//---------------------------------------------------------------------------------------------------------------
//
//  HAUD 2026.11.07
//
//  - TowerControl - fb_DisposableHeros
//
//    - this class is nothing more than the handshake sequence and a timer
//
//    - the station bitmask is written for each production cycle
//      - ticketing involves a DistributorByTicket and its companion ProcessByTicket
//      - this mock up takes care of both tickets.
//        - Why do you need to send 2 tickets?
//          - Distributor and Process instance do not know each other (and this is on purpose to keep things loose and avoid thight coupling by design)
//            --> sending tickets should be done from one place only, so a Distributor sending a ticket internally to its Process would break that rule.
//            --> The Ticket transports the information about where the movers were sent to
//              --> The Process now needs to be told which stations to activate, the rest is ruled by the bitmask from the ticket. 
//
//    - top level transport abstractions are handshaked here:
//    --------------------------------------------
//    - top level transport abstractions
//      - Instances contain the required transport logic
//      - Instances control their assigned ProcessCollector
//      - Instances are controlled in timer based application
//
//
//---------------------------------------------------------------------------------------------------------------
FUNCTION_BLOCK fb_DisposableHeros // Soldier boy, made of clay, now an empty shell
VAR_INPUT
  Start         : BOOL;           // Back to the front
  DwellTime     : TIME;           // Sounding of the clock that ticks
  StationMask   : T_PROCESS;      // molded day by day
END_VAR
VAR
  // process index
  _nProcess               : E_INSTANCE; // whoami
  _nProcessConnect        : e_instance; // to whom am I connected? this is an idea to manage the two tickets for Distributor and Process
  _nProcessConnectTarget  : e_instance; // what is the target of the process to whom I am connected

  _stInstanceCtrl         : REFERENCE TO ARRAY[1..MAX_PROCESS] OF ST_INSTANCE_CTRL;
  _stInstanceState        : REFERENCE TO ARRAY[1..MAX_PROCESS] OF ST_INSTANCE_STATE;

  _wActivateStation       : T_PROCESS;
  _stProcessData          : ST_PROCESS_DATA;

  _ItfTicketList          : I_Process_LinkedList;
  _WriteResult            : ST_PROCESS_LIST_RESULT;

  _nState                 : UINT;
  _tonProcess             : Tc2_Standard.TON;

  _nTicketCount           : UDINT;  // since this is a mock up, there is no-one to clean this up
  _nTicketCountLimit      : UDINT;  // if <> 0 --> limit is active

  _tdx                    : UINT;
END_VAR

//---------------------------------------------------------------------------------------------------------------
//---------------------------------------------------------------------------------------------------------------
// CHECK() ??
// !! this is mock up code, there is no check
//
//---------------------------------------------------------------------------------------------------------------
//---------------------------------------------------------------------------------------------------------------
IF NOT Start THEN _nState   := 0; END_IF
//---------------------------------------------------------------------------------------------------------------
CASE _nState OF
  0:
    IF Start
    THEN
      _nState               := 10;
    END_IF

  10:
    CASE _stInstanceState[_nProcess].ProcessState
    OF
      E_INSTANCE_STATE.DISABLED:
        _stInstanceCtrl[_nProcess].Cmd        := E_INSTANCE_CMD.ENABLE;
        IF (_nProcessConnect > e_instance.INSTANCE_NULL)
        THEN
          memset(ADR(_stProcessData), 0, SIZEOF(_stProcessData));
          _nState                             := 20;
          _wActivateStation                   := StationMask; // this one is important, must be double checked before sending
        END_IF

      E_INSTANCE_STATE.ENABLED:
        CASE _stInstanceState[_nProcess].ProcessProgress
        OF
          E_PROGRESS.PROGRESS_OCCUPIED:       // allow infeed movement
            _tonProcess(IN := FALSE, 
                        PT := DwellTime);

            _stInstanceCtrl[_nProcess].Cmd    := E_INSTANCE_CMD.PROCEED;
        END_CASE

      E_INSTANCE_STATE.WORKING:               // this is for the ProcessByTicket standstill handshake
        CASE _stInstanceState[_nProcess].ProcessProgress
        OF
          E_PROGRESS.PROGRESS_BUSY:           // now every mover has arrived.
            _tonProcess(IN := TRUE, 
                        PT := DwellTime);

            IF (_tonProcess.Q)
            THEN
              memset(ADR(_stProcessData), 0, SIZEOF(_stProcessData));
              _stInstanceCtrl[_nProcess].Cmd := E_INSTANCE_CMD.WORK;
            END_IF

          E_PROGRESS.PROGRESS_OCCUPIED:       // time is fleeting
            _stInstanceCtrl[_nProcess].Cmd  := E_INSTANCE_CMD.FINISH;
        END_CASE

      E_INSTANCE_STATE.FINISH:                // madness takes its toll
        CASE _stInstanceState[_nProcess].ProcessProgress
        OF
          E_PROGRESS.PROGRESS_DONE:
            _tonProcess(IN := FALSE, 
                        PT := DwellTime);

            _stInstanceCtrl[_nProcess].Cmd    := E_INSTANCE_CMD.DISABLE;

            IF (_nProcessConnect > e_instance.INSTANCE_NULL)
            THEN
              memset(ADR(_stProcessData), 0, SIZEOF(_stProcessData));
              _nState                         := 30;
              _wActivateStation               := StationMask; // this one is important, must be double checked before sending
            END_IF
        END_CASE
    END_CASE
END_CASE
CASE _nState OF
  20:
    _nState                                   :=  10;
    TruncMask();

  30:
    _nState                                   := 100;
    TruncMask();
END_CASE
CASE _nState OF

  100:
    //-----------------------------------------------------------------------------  
    // the tickets
    //-----------------------------------------------------------------------------
    // first send the ticket to the Distributor
    _WriteResult                          := _ItfTicketList.AddTailValue(_stProcessData);
    // second write the ticket for the Process
    _stProcessData.nProcessId             := _nProcessConnect;
    _stProcessData.nTargetId              := _nProcessConnectTarget;
    // third send the ticket to the Process
    _WriteResult                          := _ItfTicketList.AddTailValue(_stProcessData);
    //-----------------------------------------------------------------------------
    _nTicketCount                         := _nTicketCount + 1;;
    //-----------------------------------------------------------------------------
    _nState                               := 1000;
END_CASE
CASE _nState OF

  1000:
    IF NOT (_nTicketCountLimit > 0)
    THEN
      _nState                             := 0;
    ELSE
      IF (_nTicketCount < _nTicketCountLimit)
      THEN
        _nState                           := 0;
      END_IF
    END_IF
END_CASE

METHOD PUBLIC BitGet : BOOL
VAR_INPUT
  inVal   : T_PROCESS;
  bitNo   : DINT;
END_VAR
VAR
  wConst : T_PROCESS := 1;
END_VAR
IF ( inVal AND SHL( wConst,TO_SINT(bitNo) MOD TO_INT(SIZEOF(T_PROCESS)*8) ) ) > 0
THEN
  BitGet := TRUE;
ELSE
  BitGet := FALSE;
END_IF
END_METHOD

METHOD PUBLIC BitSet : T_PROCESS
VAR_INPUT
  inVal   : T_PROCESS;
  bitNo   : DINT;
END_VAR
VAR
  wConst  : T_PROCESS := 1;
END_VAR
BitSet := inVal OR SHL( wConst,TO_SINT(bitNo) MOD TO_INT(SIZEOF(T_PROCESS)*8) );
END_METHOD

PROPERTY InstanceCtrl : REFERENCE TO ARRAY[1..MAX_PROCESS] OF ST_INSTANCE_CTRL
SET
_stInstanceCtrl ref= InstanceCtrl;
END_SET
END_PROPERTY

PROPERTY InstanceState : REFERENCE TO ARRAY[1..MAX_PROCESS] OF ST_INSTANCE_STATE
SET
_stInstanceState ref= InstanceState;
END_SET
END_PROPERTY

PROPERTY ProcessId : E_INSTANCE
GET
ProcessId := _nProcess;
END_GET
SET
_nProcess := ProcessId;
END_SET
END_PROPERTY

PROPERTY ProcessId_Connect : E_INSTANCE
GET
ProcessId_Connect := _nProcessConnect;
END_GET
SET
_nProcessConnect := ProcessId_Connect;
END_SET
END_PROPERTY

PROPERTY ProcessId_ConnectTarget : E_INSTANCE
GET
ProcessId_ConnectTarget := _nProcessConnectTarget;
END_GET
SET
_nProcessConnectTarget := ProcessId_ConnectTarget;
END_SET
END_PROPERTY

PROPERTY TicketLinkedList : I_Process_LinkedList
SET
_ItfTicketList := TicketLinkedList;
END_SET
END_PROPERTY

METHOD TruncMask : BOOL
VAR_INPUT
END_VAR
// transfer station mask only in the range possible to handle in connected process (StationCount)
_stProcessData.nProcessId                 := _nProcess;
_stProcessData.nTargetId                  := _nProcessConnect;

FOR _tdx := 1 TO _stInstanceState[_nProcessConnect].StationCount
DO
  IF (BitGet(_wActivateStation, _tdx-1))
  THEN
    _stProcessData.wTarget                := BitSet(_stProcessData.wTarget, _tdx-1);
  END_IF      
END_FOR

TruncMask := TRUE;
END_METHOD

END_FUNCTION_BLOCK

(* stored: Version 1.1.0.1
   POU fb_DisposableHeros: Id {57ff81e0-db35-4988-adb1-755f5d46de47}, SpecialFunc None
   Method BitGet: Id {57c98de9-b3fd-4f7e-920b-502f6210a0a0}
   Method BitSet: Id {075d513b-2170-4aca-a2e9-2a16152dac6f}
   Property InstanceCtrl: Id {3363ce1e-638f-4a56-a7d9-502d7b3ac384}
   Set Set: Id {f01b16e3-e7c7-4d66-96b7-a5ce7482bb16}
   Property InstanceState: Id {4aad0611-ac13-4ac9-9913-e5032aa8988a}
   Set Set: Id {d6f80117-bb3a-400d-a886-057ce4f9cae4}
   Property ProcessId: Id {b0d1a924-6241-4335-be39-966d3f9b0719}
   Get Get: Id {4b563e78-35ca-46fa-a429-91bad99e170e}
   Set Set: Id {566aa5ef-d2c9-4a5c-8d5d-3fca3942f3dd}
   Property ProcessId_Connect: Id {abcc06e1-efe7-4aa9-9516-be1588519f38}
   Get Get: Id {b63ddabd-1e94-4d54-b9cd-0e5cfc49b660}
   Set Set: Id {97104ab0-4bc8-47e4-aa6e-413c64ff8466}
   Property ProcessId_ConnectTarget: Id {da385cf2-47a3-4307-bcdb-9af574222ed1}
   Get Get: Id {e9f241da-b82b-4801-b1f0-50eb7bef7352}
   Set Set: Id {95ea77ba-8c13-4f5b-b98e-17a763290a3b}
   Property TicketLinkedList: Id {47e1ba62-2d3b-414e-8705-080e812d120b}
   Set Set: Id {567f8792-66d5-433e-904b-9d5e5e8f13f8}
   Method TruncMask: Id {1e1b7bd6-e3e6-45f2-a35b-d0a434ac7ca6} *)
